(* IEC 61131-3 sources: Gen-AI/final/Gen-AI_v1.0_submission/A2_框架源码/agent/logs/full34_fixture/E3_P16_1_42/tools/candidate_1/fixture_compile, 1 file *)

(* ---- source.st ---- *)
FUNCTION_BLOCK FB_P16
VAR_INPUT
    processLength : USINT;
    sensor1 : BOOL;
    sensor2 : BOOL;
    sensor3 : BOOL;
    sensor4 : BOOL;
    sensor5 : BOOL;
    station1Start : BOOL;
    station2Complete : BOOL;
    station3Complete : BOOL;
    station4Complete : BOOL;
    processSequence : ARRAY[1..8] OF USINT;
END_VAR
VAR_OUTPUT
    conveyorLeft : BOOL;
    conveyorRight : BOOL;
END_VAR
(* Add a VAR block for internal state/timers before the implementation, if needed. *)
(* SKELETON ONLY: replace this RETURN with scan logic and required initial state. *)
RETURN;
END_FUNCTION_BLOCK

(* FIXTURE_COMPILE_FAIL *)
